RESOURCE RES0 : EMB_RES_ECO
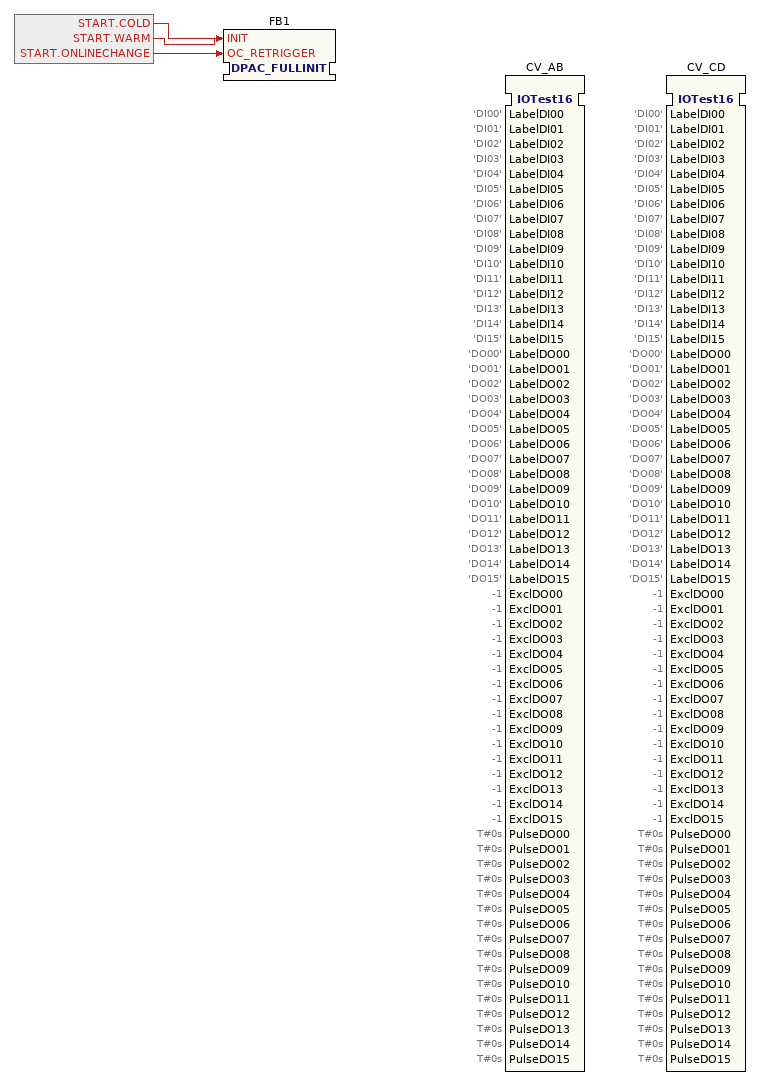
  FBS
    FB1 : DPAC_FULLINIT;
    CV_AB : IOTest16(LabelDI00 := 'DI00', LabelDO00 := 'DO00', ExclDO00 := -1, PulseDO00 := T#0s, LabelDI01 := 'DI01', LabelDO01 := 'DO01', ExclDO01 := -1, PulseDO01 := T#0s, LabelDI02 := 'DI02', LabelDO02 := 'DO02', ExclDO02 := -1, PulseDO02 := T#0s, LabelDI03 := 'DI03', LabelDO03 := 'DO03', ExclDO03 := -1, PulseDO03 := T#0s, LabelDI04 := 'DI04', LabelDO04 := 'DO04', ExclDO04 := -1, PulseDO04 := T#0s, LabelDI05 := 'DI05', LabelDO05 := 'DO05', ExclDO05 := -1, PulseDO05 := T#0s, LabelDI06 := 'DI06', LabelDO06 := 'DO06', ExclDO06 := -1, PulseDO06 := T#0s, LabelDI07 := 'DI07', LabelDO07 := 'DO07', ExclDO07 := -1, PulseDO07 := T#0s, LabelDI08 := 'DI08', LabelDO08 := 'DO08', ExclDO08 := -1, PulseDO08 := T#0s, LabelDI09 := 'DI09', LabelDO09 := 'DO09', ExclDO09 := -1, PulseDO09 := T#0s, LabelDI10 := 'DI10', LabelDO10 := 'DO10', ExclDO10 := -1, PulseDO10 := T#0s, LabelDI11 := 'DI11', LabelDO11 := 'DO11', ExclDO11 := -1, PulseDO11 := T#0s, LabelDI12 := 'DI12', LabelDO12 := 'DO12', ExclDO12 := -1, PulseDO12 := T#0s, LabelDI13 := 'DI13', LabelDO13 := 'DO13', ExclDO13 := -1, PulseDO13 := T#0s, LabelDI14 := 'DI14', LabelDO14 := 'DO14', ExclDO14 := -1, PulseDO14 := T#0s, LabelDI15 := 'DI15', LabelDO15 := 'DO15', ExclDO15 := -1, PulseDO15 := T#0s);
    CV_CD : IOTest16(LabelDI00 := 'DI00', LabelDO00 := 'DO00', ExclDO00 := -1, PulseDO00 := T#0s, LabelDI01 := 'DI01', LabelDO01 := 'DO01', ExclDO01 := -1, PulseDO01 := T#0s, LabelDI02 := 'DI02', LabelDO02 := 'DO02', ExclDO02 := -1, PulseDO02 := T#0s, LabelDI03 := 'DI03', LabelDO03 := 'DO03', ExclDO03 := -1, PulseDO03 := T#0s, LabelDI04 := 'DI04', LabelDO04 := 'DO04', ExclDO04 := -1, PulseDO04 := T#0s, LabelDI05 := 'DI05', LabelDO05 := 'DO05', ExclDO05 := -1, PulseDO05 := T#0s, LabelDI06 := 'DI06', LabelDO06 := 'DO06', ExclDO06 := -1, PulseDO06 := T#0s, LabelDI07 := 'DI07', LabelDO07 := 'DO07', ExclDO07 := -1, PulseDO07 := T#0s, LabelDI08 := 'DI08', LabelDO08 := 'DO08', ExclDO08 := -1, PulseDO08 := T#0s, LabelDI09 := 'DI09', LabelDO09 := 'DO09', ExclDO09 := -1, PulseDO09 := T#0s, LabelDI10 := 'DI10', LabelDO10 := 'DO10', ExclDO10 := -1, PulseDO10 := T#0s, LabelDI11 := 'DI11', LabelDO11 := 'DO11', ExclDO11 := -1, PulseDO11 := T#0s, LabelDI12 := 'DI12', LabelDO12 := 'DO12', ExclDO12 := -1, PulseDO12 := T#0s, LabelDI13 := 'DI13', LabelDO13 := 'DO13', ExclDO13 := -1, PulseDO13 := T#0s, LabelDI14 := 'DI14', LabelDO14 := 'DO14', ExclDO14 := -1, PulseDO14 := T#0s, LabelDI15 := 'DI15', LabelDO15 := 'DO15', ExclDO15 := -1, PulseDO15 := T#0s);
  END_FBS
  EVENT_CONNECTIONS
    START.COLD TO FB1.INIT;
    START.WARM TO FB1.INIT;
    START.ONLINECHANGE TO FB1.OC_RETRIGGER;
  END_CONNECTIONS
END_RESOURCE
